(* IEC 61131-3 sources: 2026_Projet_YGO_ExcavatriceDragage/CODE/J_SUPERVISION/_TYPES/6_DIAG_ET_CHAINES, 10 files *)

(* ---- ST_ChainContextGlobal.st ---- *)
TYPE ST_ChainContextGlobal :
STRUCT
    Idx101_ModeActive             : E_Mode; // Mode de marche actif (MANUEL, SEMI_AUTO, MAINT_N1, MAINT_N2)
    Idx102_SimulationEnabled      : BOOL;   // 0 = Matériel Réel (Nominal) | 1 = SIMULATION ACTIVE ⚠️
    Idx103_JoystickCommOk         : BOOL;   // 1 = Comm CANopen Joystick OK (Sain) | 0 = Perte Comm CAN

    Idx201_JoystickSelected       : BOOL;   // 1 = Pilotage par Joystick Hall | 0 = Pilotage par Boutons IHM
    Idx202_BypassNetworkGlobal    : BOOL;   // 0 = Comm Réseau OK | 1 = BYPASS RÉSEAU ACTIF ⚠️
    Idx203_BypassSensorsGlobal    : BOOL;   // 0 = Capteurs Actifs | 1 = AU MOINS 1 CAPTEUR SHUNTÉ ⚠️

    Idx301_EmergencyChainClosed   : BOOL;   // 1 = Boucle AU Matérielle Fermée (OK) | 0 = AU APPUYÉ
    Idx302_PowerContactorEngaged  : BOOL;   // 1 = Puissance Armée | 0 = Puissance Coupée
    Idx303_SafeStopActiveAny      : BOOL;   // 0 = Sain | 1 = AU MOINS UN SAFESTOP MÉTIER ACTIF
    Idx304_PowerCutOffActiveAny   : BOOL;   // 0 = Sain | 1 = COUPURE GENERAL COLLAGE ACTIVEE

    Idx401_HmiHeartbeatOk         : BOOL;   // 1 = Liaison IHM Active | 0 = Perte Liaison IHM
    Idx402_CycleAutoBusy          : BOOL;   // 1 = Séquenceur Auto en Cours | 0 = Repos
END_STRUCT
END_TYPE

(* ---- ST_EmergencyCmd.st ---- *)
(* ═══════════════════════════════════════════════════════════════
   🎮 ST_EmergencyCmd — Commandes IHM de la chaîne AU / sécurité
   ───────────────────────────────────────────────────────────────
   🎯 Rôle : Commandes opérateur (boutons IHM) de la chaîne d'arrêt
      d'urgence, sorties de `Modes.Cmd`. Point de vue IHM : `Cmd` =
      les boutons. Distinctes des commandes physiques fail-safe
      `ST_Safety_Emergency_Cmd` (MaintainA/B_Cmd, ArmPulse_Cmd) qui
      sont des sorties du FB AU, internes à PRG_06 — PAS des commandes
      IHM.
   🔌 Interface : Produit par l'IHM, consommé par PRG_02 / PRG_06 /
      FB_TroubleshootingView.
   📄 Doc : DOC/AF/AF_Partie-01_Analyse_Fonctionnelle_v2.1.md §5
   ═══════════════════════════════════════════════════════════════ *)
TYPE ST_EmergencyCmd :
STRUCT
    BtnEmergencyArming : BOOL;   (* 🎮 Commande IHM réarmement contacteur puissance (front) — PAS de réarmement automatique *)
    BtnEmergencyCutOff : BOOL;   (* 🎮 Commande IHM coupure d'urgence puissance amont (arrêt à distance) *)
END_STRUCT
END_TYPE

(* ---- ST_EmergencyHMI.st ---- *)
(* ═══════════════════════════════════════════════════════════════
   🛡️ ST_EmergencyHMI — Données d'échange IHM de la chaîne AU / sécurité
   ───────────────────────────────────────────────────────────────
   🎯 Rôle : Structure dédiée `GVL_IHM.Emergency`. Regroupe les
      champs emergency/safety sortis de `Modes`, selon le standard IHM
      projet (Cmd + State [+ Cfg]) :
        • Cmd   : ST_EmergencyCmd              (boutons opérateur IHM)
        • State : ST_EmergencyState            (état AU + cmd FB AU + Diag interne)
      Point de vue IHM : `Cmd` = les boutons. Les commandes physiques
      fail-safe (MaintainA/B_Cmd, ArmPulse_Cmd) sont des sorties du FB
      AU, exposées dans `State` comme states/info. Le diagnostic vit
      dans `State.Diag` (PAS de dossier `Diag` au top).
   🔌 Interface : Produit par PRG_07_Supervision (State) et
      l'IHM (Cmd), consommé par PRG_02 / PRG_06 / FB_TroubleshootingView.
   📄 Doc : DOC/AF/AF_Partie-01_Analyse_Fonctionnelle_v2.1.md §5
   ═══════════════════════════════════════════════════════════════ *)
TYPE ST_EmergencyHMI :
STRUCT
    Cmd   : ST_EmergencyCmd;   // 🎮 Boutons opérateur IHM (réarmement / coupure)
    State : ST_EmergencyState; // 📊 État AU + cmd FB AU + Diag interne
END_STRUCT
END_TYPE

(* ---- ST_EmergencyState.st ---- *)
(* ═══════════════════════════════════════════════════════════════
   📊 ST_EmergencyState — État IHM de la chaîne AU / sécurité
   ───────────────────────────────────────────────────────────────
   🎯 Rôle : État/diagnostic IHM de la chaîne d'arrêt d'urgence,
      sorti de `Modes.State`. Point de vue IHM : `State` regroupe les
      champs d'état AU (ChainOk, ContactorOk, Armable, ArmingBusy, Step)
      en champs plats, les commandes physiques fail-safe du FB AU
      (MaintainA/B_Cmd, ArmPulse_Cmd) exposées comme states/info, et le
      diagnostic AU (`Diag : ST_Safety_Emergency_Diag`) en structure
      interne. PAS de sous-State imbriqué, PAS de dossier `Diag` au top
      de `Emergency` — le diagnostic vit dans `State`.
   🔌 Interface : Produit par PRG_07_Supervision, consommé par l'IHM.
   📄 Doc : DOC/AF/AF_Partie-01_Analyse_Fonctionnelle_v2.1.md §5
   ═══════════════════════════════════════════════════════════════ *)
TYPE ST_EmergencyState :
STRUCT
    // ── État AU (champs plats, miroir du DUT AU ST_Safety_Emergency_State) ──
    ChainOk     : BOOL; // Boucle AU fermee (EmergencyChainClosed = TRUE)
    ContactorOk : BOOL; // Contacteur puissance confirme engage (PowerContactorEngaged = TRUE)
    Step        : INT;  // Etape sequence armement : 0=IDLE, 1=TestA, 2=RestoreA, 3=TestB, 4=RestoreB, 5=Pulse, 6=Confirm
    Armable     : BOOL; // Rearmement possible maintenant : chain OK, step=0, pas de lockout
    ArmingBusy  : BOOL; // Sequence armement OU lockout en cours (nouvelle demande ignoree)

    // ── États publics FB AU (Ready/Done/Fault/OperatorMessage) ──
    // Miroir des champs Status du FB_Safety_EmergencyManagement (produits par PRG_06).
    // Busy n'est PAS exposé : redondant avec ArmingBusy (déjà présent ci-dessus).
    Ready           : BOOL; // FB AU pret a fonctionner (Enable + pas de StartupFail)
    Done            : BOOL; // Cycle rearmement AU termine (contacteur puissance confirme engage)
    Fault           : ST_Fault; // Defaut latte de la chaine AU (socle FB_FaultCore, vue live + latchee)
    OperatorMessage : STRING(120); // Message operateur par etat / par probleme de la chaine AU

    // ── Commandes physiques fail-safe du FB AU (exposées comme states/info) ──
    MaintainA_Cmd : BOOL; // Sortie pilotage canal A (TRUE = voie maintenue) — interne FB AU
    MaintainB_Cmd : BOOL; // Sortie pilotage canal B (TRUE = voie maintenue) — interne FB AU
    ArmPulse_Cmd  : BOOL; // Impulsion rearmement physique (1s) — interne FB AU

    // ── Diagnostic AU (structure interne de State) ──
    Diag : ST_Safety_Emergency_Diag; // Diagnostic et erreurs de la chaîne AU
END_STRUCT
END_TYPE

(* ---- ST_HomingChecklist.st ---- *)
(* ═══════════════════════════════════════════════════════════════
   🎯 ST_HomingChecklist — Diagnostic chronologique de référencement (Dépannage)
   ───────────────────────────────────────────────────────────────
   🎨 Permet de localiser immédiatement l'étape qui bloque le Homing (M1/M2).
   ═══════════════════════════════════════════════════════════════ *)
TYPE ST_HomingChecklist :
STRUCT
    (* 1. Pré-requis de mode *)
    Step1_ModeAuthorized         : BOOL; (* TRUE = Mode MAINT_N1 ou MAINT_N2 actif ➔ Commutateur Mode IHM : GVL_IHM.Modes *)
    Step2_WinchSelected          : BOOL; (* TRUE = Treuil sélectionné en MAINT_N2 ➔ Bouton IHM : GVL_IHM.Modes.Cmd.TglJoystickMaster / Selection Treuil *)

    (* 2. Santé Matériel & Bus *)
    Step3_EncoderAvailable       : BOOL; (* TRUE = Codeur EtherCAT OK & E/S OK ➔ Si simu : GVL_Simulation.SimWinchActive=1 / SimSafetyActive=1 *)

    (* 2bis. Entrées physiques directes HwIn (vérité terrain) *)
    HwIn_ContactorsReleased_DI   : BOOL; (* Retours contacteurs retombés issus de HwIn.Winch *)
    HwIn_BrakeIsOpen_DI          : BOOL; (* Retour fin de course frein (1 = ouvert) issu de HwIn.Winch *)
    HwIn_TopPositionFree_DI      : BOOL; (* Capteur position haute commun libre (1 = libre) issu de HwIn.Winch *)

    (* 3. État Physique Machine *)
    Step4_ContactorsReleased     : BOOL; (* TRUE = Tous les contacteurs retombés (attendre l'arrêt complet) *)
    Step5_BrakeApplied           : BOOL; (* TRUE = Frein serré (attendre l'arrêt complet) *)
    TopPositionSensorActive      : BOOL; (* 📍 Fin de course haut physique (TRUE = au contact) *)
    BucketIsOpen                 : BOOL; (* 🪣 Benne Ouvert (TRUE = Ouvert) ➔ Pour forcer sans codeur : GVL_IHM.M2TreuilBenne.Bucket.Cmd.BtnConfirmOpenPos *)

    (* 4. Séquence & Bilan *)
    AllConditionsMet             : BOOL; (* TRUE = Prêt pour le homing ! ➔ Déclencher : GVL_IHM.M1TreuilRetenue.Cmd.BtnHome (à 8m) ou BtnHomingAtZero (à 0m) *)
    HomingBusy                   : BOOL; (* TRUE = Séquence de calage en cours *)
    HomingDone                   : BOOL; (* TRUE = Calage réussi *)
    HomingHomed                  : BOOL; (* TRUE = Treuil actuellement référencé *)
    HomingSuspect                : BOOL; (* TRUE = Doute redémarrage ➔ Lever le doute via : GVL_IHM.M1TreuilRetenue.Cmd.BtnConfirmCoherence *)

    (* 5. Code de rejet exact *)
    RejectErrorMask              : WORD; (* Bitmask d'erreur FB_Encoder_Homing.ErrorId *)
    TopContactLatched            : BOOL; (* Contact TOP touche pendant cycle homing (degagement en cours) *)
    TopContactCount              : UINT; (* Compteur contacts capteur TOP pendant cycle homing *)
END_STRUCT
END_TYPE

(* ---- ST_InputModuleDiagHMI.st ---- *)
(* ═══════════════════════════════════════════════════════════════
   🩺 ST_InputModuleDiagHMI — Diagnostic carte des modules DI TOR réelles
   ───────────────────────────────────────────────────────────────
   📄 Doc métier : DOC/AF/AF_Partie-06_Acquisition_Qualification_IO_v2.4.md §3bis
   🎨 Granularité MODULE (pas canal) : GetDeviceState() est un état de carte,
      pas un diagnostic par voie. Un module en défaut ne dit pas *quelle*
      TOR ment, seulement qu'aucune des TOR qu'il porte n'est fiable.
   🔗 Producteur : PRG_02_Acquisition (3 appels GetDeviceState()).
   ═══════════════════════════════════════════════════════════════ *)
TYPE ST_InputModuleDiagHMI :
STRUCT
    LocalDigitalIoOk : BOOL; (* TRUE = module Local_Digital_IO opérationnel (8 TOR Winch/Machine) *)
    Vh0800EndOk      : BOOL; (* TRUE = module VH_0800END opérationnel (7 TOR freins/thermiques/AU) *)
    Vh0808EtpOk      : BOOL; (* TRUE = module VH_0808ETP opérationnel (7 TOR positions M3/hydraulique/crible) *)
    Vh0008ErOk       : BOOL; (* TRUE = module VH_0008ER opérationnel (8 DO Relais Freins/Kobold) *)
    Vh0008Er1Ok      : BOOL; (* TRUE = module VH_0008ER_1 opérationnel (8 DO Relais AU/PowerKeepAlive) *)
    Fault            : BOOL; (* TRUE = au moins un des 5 modules E/S hors service *)
END_STRUCT
END_TYPE

(* ---- ST_IOModuleDiag.st ---- *)
(* ═══════════════════════════════════════════════════════════════
   🩺 ST_IOModuleDiag — Diagnostic carte des 5 modules E/S physiques
   ───────────────────────────────────────────────────────────────
   📄 Doc métier : DOC/AF/AF_Partie-06_Acquisition_Qualification_IO_v2.4.md §3bis
   🎨 Granularité MODULE (pas canal) : GetDeviceState() est un état de carte,
      pas un diagnostic par voie. Un module en défaut ne dit pas *quelle*
      TOR ment, seulement qu'aucune des TOR qu'il porte n'est fiable.
   🔗 Producteur : PRG_02_Acquisition (5 appels GetDeviceState()).
   🔌 Consommateurs : PRG_04 (SafeStop treuils), PRG_05 (SafeStop M3),
      PRG_07 (recopie IHM GVL_IHM.Network.InputModules + FB_TroubleshootingView).
   ═══════════════════════════════════════════════════════════════ *)
TYPE ST_IOModuleDiag :
STRUCT
    LocalDigitalIoOk : BOOL;  // Module Local_Digital_IO OK (DI8/DO8)
    Vh0800EndOk      : BOOL;  // Module VH_0800END OK (DI8)
    Vh0808EtpOk      : BOOL;  // Module VH_0808ETP OK (DI8/DO8)
    Vh0008ErOk       : BOOL;  // Module VH_0008ER OK (DO8 Relais Freins/Kobold)
    Vh0008Er1Ok      : BOOL;  // Module VH_0008ER_1 OK (DO8 Relais AU/PowerKeepAlive)
    Fault            : BOOL;  // Défaut sur au moins un module E/S
END_STRUCT
END_TYPE

(* ---- ST_MotionChecklist.st ---- *)
(* ═══════════════════════════════════════════════════════════════
   ⚙️ ST_MotionChecklist — Diagnostic chronologique de commande de mouvement
   ───────────────────────────────────────────────────────────────
   🎨 Permet de voir en un coup d'œil pourquoi un ordre de mouvement ne fait pas coller les relais.
   ═══════════════════════════════════════════════════════════════ *)
TYPE ST_MotionChecklist :
STRUCT
    (* 1. Puissance & Mode *)
    Step1_PowerEngaged           : BOOL; (* TRUE = Contacteur principal sous tension (PowerContactorEngaged_DI) ➔ Armer puissance via Reset *)
    Step2_ModeAuthorized         : BOOL; (* TRUE = Mode MAINT_N1 ou N2 actif (pas DISABLE) ➔ Commutateur Mode IHM *)
    Step3_NotBusyOtherTask       : BOOL; (* TRUE = Pas d'autre séquence en cours (Homing, Benne busy, etc.) *)

    (* 1bis. Entrées physiques directes HwIn (vérité terrain) *)
    HwIn_PowerContactorEngaged_DI: BOOL; (* Contacteur puissance principal issu de HwIn.Machine *)
    HwIn_BrakeIsOpen_DI          : BOOL; (* Retour fin de course frein (1 = ouvert) issu de HwIn *)
    Cmd_BrakeRelease             : BOOL; (* Ordre de commande d'ouverture de frein généré par l'automate *)

    (* 2. Intention & Demande *)
    Step4_MotionRequested        : BOOL; (* TRUE = Demande active (Bouton IHM ou Joystick) ➔ Si IHM : TglJoystickMaster doit être à 0 ! *)
    RequestedDirection           : INT;  (* +1 = Ascending, -1 = Descending, 0 = Repos *)
    RequestedSpeedPct            : REAL; (* 0..100 % consigne demandée *)

    (* 3. Chaîne de Sécurité & Verrous *)
    Step5_NoSafetyFault          : BOOL; (* TRUE = Pas de SafeStop ni AU actif sur cet axe *)
    Step6_DirectionAllowed       : BOOL; (* TRUE = Sens autorisé (AscentPermit/DescendPermit / TremiePermit/MaintenancePermit) *)
    Step7_BrakeReleased          : BOOL; (* TRUE = Commande frein activée & retour frein OK *)
    Step8_OutputInterlockOk      : BOOL; (* TRUE = Étage de sortie LD débloqué (pas d'interlock actif).
                                             🛡️ T371 : dérivé de l'ÉTAT publié + du défaut de la barrière finale,
                                             JAMAIS du seul FinalInterlockError (qui ne porte que le timeout frein). *)

    (* 4. Bilan & Exécution Physiques *)
    AllConditionsMet             : BOOL; (* 🟢 TRUE = TOUTES LES CONDITIONS SONT REMPLIES, LES RELAIS DOIVENT COLLER ! *)
    RelayFwdActive               : BOOL; (* 🛗 Relais Ascending physiquement commandé *)
    RelayRevActive               : BOOL; (* 🛗 Relais Descending physiquement commandé *)
    SpeedContactor1Active        : BOOL; (* 🔌 Contacteur de vitesse Palier 1 commandé *)

    (* 5. Barrière finale — état & cause publiés (T371, LECTURE SEULE) *)
    (* ⚠️ Ajout en FIN de STRUCT : aucun champ existant n'est décalé (mapping IHM/SCADA + online change).
       ⚠️ VOCABULAIRE COMMUN aux 3 axes (famille E_WinchFinalInterlock...), choisi parce que ce DUT est
          PARTAGÉ par M1, M2 et M3 et qu'AUCUNE conversion de type n'est nécessaire :
          · M1/M2 — recopie DIRECTE de l'énumération publiée par la barrière (aucune projection) ;
          · M3   — la barrière M3 ne publie qu'un état dérivé du défaut : E_State.READY -> READY et
                   E_State.ERROR -> FAULT (projection EXPLICITE, cf. FB_TroubleshootingView.st §11),
                   ses 3 raisons étant identiques (NONE / BRAKE_COMMAND_NOT_CONFIRMED / RESTART_INHIBITED).
          Le type énuméré (et non INT) évite toute conversion — la conversion explicite de l'énumération
          d'un membre d'IEC_STRUCT n'est pas supportée par le compilateur de test, et un INT aurait rendu
          la table de valeurs DÉPENDANTE DE L'AXE. La famille M3 (E_State) n'est volontairement pas
          réutilisée ici : sa numérotation diffère (READY = 2 vs 1) et rendrait la lecture ambiguë.
       ⚠️ USAGE DIAGNOSTIC UNIQUEMENT (latence N-1 assumée, projection PRG_04:1688-1696) : aucune ligne
          de CONDUITE ne doit consommer ces deux champs. *)
    Step8_InterlockState         : E_WinchFinalInterlockState;  (* 🛡️ [DIAG/LECTURE] État publié de la barrière
                                             finale, vocabulaire commun aux 3 axes :
                                             DISABLED(0) · READY(1) · WAIT_BRAKE_COMMAND_CONFIRMATION(2) ·
                                             WAIT_STEP_DELAY(3) · WAIT_RESTART_DELAY(4) · FAULT(5) ·
                                             WAIT_SENSE_DROP_CONFIRM(6).
                                             ⚠️ WAIT_STEP_DELAY(3) n'est JAMAIS produit : `FB_WinchOutputInterlock.st`
                                                ne l'affecte nulle part (la montée de palier reste en READY, :473) —
                                                entrée conservée pour la complétude de l'énumération (REX revue T371). *)
    Step8_InterlockReason        : E_WinchFinalInterlockReason; (* 🛡️ [DIAG/LECTURE] Cause MÉMORISÉE publiée par la
                                             barrière finale, vocabulaire commun aux 3 axes :
                                             NONE(0) · BRAKE_COMMAND_NOT_CONFIRMED(1) · RESTART_INHIBITED(2) ·
                                             SENSE_DROP_TIMEOUT(3 — M1/M2 uniquement).
                                             ⚠️ Cause mémorisée, JAMAIS remise à NONE par un acquittement sur
                                                certains chemins (SENSE_DROP_TIMEOUT M1/M2, RESTART_INHIBITED M3) :
                                                elle informe, elle ne prouve pas un refus ACTIF. *)
END_STRUCT
END_TYPE

(* ---- ST_NetworkDiagHMI.st ---- *)
(* ═══════════════════════════════════════════════════════════════
   📡 ST_NetworkDiagHMI — Données d'échange IHM pour les diagnostics réseau
   ───────────────────────────────────────────────────────────────
   🎨 Destiné à l'affichage des diagnostics CANopen et EtherCAT.
   ═══════════════════════════════════════════════════════════════ *)
TYPE ST_NetworkDiagHMI :
STRUCT
    BusCanOpen          : ST_Diag_Device;  (* 📡 Diagnostics bus CANopen *)
    Joystick            : ST_Diag_Device;  (* 🕹️ Diagnostics esclave Joystick *)
    CanError            : BOOL;           (* ⚠️ Voyant anomalie globale CANopen (IHM Visu) *)
    CanErrorId          : WORD;           (* ❌ Code anomalie CANopen *)

    BusEthercat         : ST_Diag_Device;  (* 📡 Diagnostics bus EtherCAT *)
    EncoderM1           : ST_Diag_Device;  (* 🧲 Diagnostics esclave COD1 *)
    EncoderM2           : ST_Diag_Device;  (* 🧲 Diagnostics esclave COD2 *)
    VariateurM3         : ST_Diag_Device;  (* ↔️ Diagnostics esclave AC600 *)
    EcatError           : BOOL;           (* ⚠️ Voyant anomalie globale EtherCAT (IHM Visu) *)
    EcatErrorId         : WORD;           (* ❌ Code anomalie EtherCAT *)

    InputModules        : ST_InputModuleDiagHMI; (* 🩺 Diagnostic carte des 5 modules d'E/S physiques *)

    (* 🌐 Bypass réseau global *)
    Bypass              : ST_BypassNetwork;
END_STRUCT
END_TYPE

(* ---- ST_SafetyChecklist.st ---- *)
(* ═══════════════════════════════════════════════════════════════
   🛡️ ST_SafetyChecklist — Diagnostic chronologique réarmement chaîne de sécurité / AU
   ───────────────────────────────────────────────────────────────
   🎨 Permet d'identifier immédiatement pourquoi la puissance / AU ne réarme pas.
   ═══════════════════════════════════════════════════════════════ *)
TYPE ST_SafetyChecklist :
STRUCT
    (* 0. Aiguillage source — dit QUELLE entree alimente les steps 1-3 ci-dessous.
       Absent jusqu'ici : diagnostiquer un blocage AU en full simu obligeait a rouvrir
       GVL_Simulation dans un Watch separe (, banc sans HW). *)
    SimulationModeActive         : BOOL; (* TRUE = bit maitre simu actif (GVL_Simulation.SimulationModeActive) *)
    SimSafetyActive              : BOOL; (* TRUE = domaine Safety simule ➔ Step1-3 lisent FB_Sim_Safety, pas les DI/comm reelles *)

    (* 0bis. Entrées physiques directes HwIn (vérité terrain) *)
    HwIn_EmergencyChainClosed_DI : BOOL; (* Boucle AU physique ou simulée issue de HwIn.Machine *)
    HwIn_PowerContactorEngaged_DI: BOOL; (* Retour contacteur de puissance issu de HwIn.Machine *)
    HwIn_EmergencyBtnCut_HMI     : BOOL; (* Commande coupure AU IHM *)

    (* 1. Intégrité matérielle & modules E/S *)
    Step1_InputModulesOk         : BOOL; (* TRUE = Les 3 cartes E/S physiques sont RUNNING ➔ En simu : GVL_Simulation.SimSafetyActive=1 *)
    Step2_EmergencyBtnNotCut     : BOOL; (* TRUE = Pas d'appui AU ➔ Déverrouiller le BP coup-de-poing physique ou IHM : GVL_IHM.Modes.Cmd.BtnEmergencyCutOff *)
    Step3_EmergencyChainClosed   : BOOL; (* TRUE = Boucle physique AU fermée (EmergencyChainClosed_DI) *)

    (* 2. Conditions de réarmement *)
    Step4_ContactorReleased      : BOOL; (* TRUE = Contacteur relâché ; précondition AF01 avant réarmement *)
    Step5_ArmingAllowed          : BOOL; (* TRUE = Armable ; acquitter si nécessaire puis générer un front BtnEmergencyArming *)

    (* 3. Séquence de réarmement *)
    ArmingStep                   : INT;  (* 0=IDLE, 1=TestA, 2=RestoreA, 3=TestB, 4=RestoreB, 5=Pulse, 6=Confirm *)
    ArmingPulseActive            : BOOL; (* TRUE = Impulsion d'armement en cours *)
    ArmingBusy                   : BOOL; (* TRUE = séquence de réarmement ou verrouillage en cours *)
    LockoutActive                : BOOL; (* TRUE = verrouillage temporel entre tentatives *)
    PowerContactorEngaged        : BOOL; (* TRUE = Contacteur principal sous tension (PowerContactorEngaged_DI) *)
    PowerCutOffActive            : BOOL; (* TRUE = demande de coupure safety active *)
    PowerCutOffRequest           : BOOL; (* TRUE = demande de coupure AU (entrée instSafetyEmergencyManagement) *)
    MaintainAActive              : BOOL; (* TRUE = maintien voie A demandé *)
    MaintainBActive              : BOOL; (* TRUE = maintien voie B demandé *)
    AllConditionsMet             : BOOL; (* TRUE = état final : chaîne OK et puissance engagée *)

    (* 4. Erreurs *)
    SafetyError                  : BOOL; (* TRUE = Défaut sécurité actif *)
    ArmingErrorId               : WORD; (* bit0 redondance ; bit1 échec confirmation contacteur *)
    RedundancyTestFailed         : BOOL; (* TRUE = Défaut test de redondance contacteurs *)
    ArmingFailed                 : BOOL; (* TRUE = Échec de la séquence d'armement *)
    WasArmed                     : BOOL; (* TRUE = AU armée au moins une fois ; PowerKeepAlive maintenu à travers un appui AU pur *)
    LastAbortStep                : INT;  (* Étape atteinte lors du dernier abandon de séquence (0..6) *)
    LastAbortCause               : WORD; (* Cause du dernier abandon (masque bitfield) *)
END_STRUCT
END_TYPE
